// TIA Portal V21 export
// export: Created 2026-11-21T13:00:31.813493Z, ExportSetting WithDefaults, DisplayName Totally Integrated Automation Portal, DisplayVersion V21, DisplayName STEP 7 Professional, DisplayVersion V21, DisplayName STEP 7 Safety, DisplayVersion V21, DisplayName Tech WebApplication, DisplayVersion V21, DisplayName WinCC Basic/Comfort/Advanced, DisplayVersion V21, DisplayName WinCC Unified, DisplayVersion V21
PlcWatchTable "Outputs"
  PlcWatchTableEntry ""Motor""  DisplayFormat=Bool, ModifyTrigger=Permanent, MonitorTrigger=Permanent
  PlcWatchTableEntry ""Alarm""  DisplayFormat=Bool, ModifyTrigger=Permanent, MonitorTrigger=PermanentAtEnd
